Fanuc KAREL source: ka00067.KL

PROGRAM KA00067
%STACKSIZE=65535
%PRIORITY=65535
%NOLOCKGROUP
VAR
SRC : XYZWPR
DST : XYZWPREXT
BEGIN
SRC.X=1.0
-- UNSAFE_SOURCE_IR line 8: DST = convert_xyzwpr_to_xyzwprext(SRC)
END KA00067
